{attribute 'qualified_only'}
{attribute 'strict'}
TYPE E_SignalQuality :
(
    Good                := 0,
    BadComm             := 1,
    BadConfig           := 2,
    BadDeviceFault      := 3,
    UncertainStale      := 4,
    UncertainInit       := 5
) UINT;
END_TYPE

(* stored: Version 1.1.0.1, ProductVersion 3.1.4024.0
   DUT E_SignalQuality: Id {182781b4-018b-4181-aae4-73847ac012ed} *)
